(* PLC project Vn_two_rungs, Beckhoff Automation GmbH TwinCAT PLC Control 3.5.13.21 *)
(* stored: creationDateTime 1970-01-01T00:00:00 *)

PROGRAM Vn_two_rungs

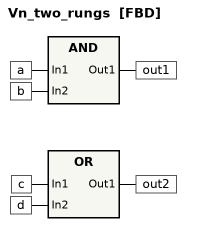
(* FBD diagram, written out as Structured Text *)
out1 := a AND b;
out2 := c OR d;
END_PROGRAM
